Fanuc KAREL source: kt00477.KL

-- PROVISIONAL review KL for V770-1; original PC SHA256 4bb35c99dc1c48e64c0b877d203e75de5b974a8a8edab8cca158433a3996d53e
-- Incomplete behavior may be omitted. Consult companion uncertainty JSON. Do not deploy.
PROGRAM KT00477
%NOLOCKGROUP
-- UNRESOLVED_DECL P1 type=000101
-- UNRESOLVED_DECL P2 type=000101
-- UNRESOLVED_DECL OUT type=000199
BEGIN
  -- UNRESOLVED_PC offsets 5-34; opcodes 49,49,60,7E,4A
  -- UNRESOLVED_PC offsets 39-43; opcodes 7F
END KT00477
